Staubli VAL3: Motion.pjx

--- Motion.pjx ---
Parameters version=s8.15.3Cs9_BS3337 stackSize=200000 millimeterUnit=true
Program file=getMoveDone.pgx
Program file=home.pgx
Program file=moveToPoint.pgx
Program file=setSpeed.pgx
Data file=Motion.dtx
Library alias=io path=Disk://io/io.pjx autoload=true password=

--- Motion.dtx ---
public mdesc mNomSpeed = {accel=25, vel=20, decel=25, blend=off, leave=0, reach=0}
public mdesc mFine = {accel=10, vel=10, decel=10, blend=off, leave=0, reach=0}
public joint jHome
public tool tTool = {fatherId=flange[0]}

--- getMoveDone.pgx ---
public program getMoveDone(num& x_nResult)
  local num l_nT0
  local num l_nTimeout
//等待已下发的运动全部执行完，并等到机械臂停稳
//返回码 x_nResult：0=已停稳  1=指令执行完但 2s 内仍未停稳（残余抖动/受外力）
//依据：waitEndMove() 手册 10.6 第177页；isSettled() 手册 10.6 第178页
begin
  x_nResult=0

  //1) 取消上一条指令的混接，并等它执行完（手册 10.6，第177页）
  //   注意：waitEndMove 只等到"位置指令下发到位"，不等机械臂稳定
  waitEndMove()

  //2) 需要完全停稳时必须再用 isSettled()（手册 10.6，第178页）
  l_nTimeout=2
  if isSettled()==false
    l_nT0=clock()                                  //手册 5 章，第103页
    do
      delay(0.01)                                  //循环里必须让出 CPU
    until (isSettled()==true) or ((clock()-l_nT0)>=l_nTimeout)
    //超时不抛错：有的工位（打磨/压装）本来就有持续微振，交给调用方判断
    if isSettled()==false
      x_nResult=1
    endIf
  endIf
end

--- home.pgx ---
public program home(num& x_nResult)
  local num l_nMoveId
//关节运动(movej)回 Home 位 jHome，并等待到位/停稳
//返回码 x_nResult：0=已到 Home 并停稳  1=到点但仍有残余抖动  -2=jHome 超出软件限位
//依赖：Motion.dtx 的 jHome（当前是全 0 占位，示教后才是真实 Home）
begin
  x_nResult=0

  waitEndMove()

  //jHome 现在是全 0 占位，先判软件限位（bool isInRange(joint)，手册 9.2，第133页）；
  //不在限位内就直接返回错误，不要让控制器抛 runtime error
  if isInRange(jHome)==false
    x_nResult=-2
    return
  endIf

  //movej 的第一个参数必须用 joint 变量传入；写成 {0,0,0,0,0,0} 会被判为歧义表达式
  //（手册 10.6，第173页 movej 的 Example 有说明）
  l_nMoveId=movej(jHome,tTool,mFine)

  //move id 只能用 >= 判断，且完成判据是 +1（手册 10.4，第180页）
  wait(getMoveId()>=l_nMoveId+1)

  call getMoveDone(x_nResult)
end

--- moveToPoint.pgx ---
public program moveToPoint(point x_pTarget, tool x_tTool, mdesc x_mDesc, num& x_nResult)
  local num l_nMoveId
//直线运动(movel)到点位，并等待到位/停稳
//用法：call mot:moveToPoint(pPick, mot:tTool, mot:mNomSpeed, nResult)
//      要精定位时把第 3 个参数换成 mot:mFine
//返回码 x_nResult：0=已到位并停稳  1=指令执行完但仍有残余抖动（见 getMoveDone）  2=运动被中断
//点位由调用方传入（本库不放占位点位，见 Motion.dtx 注释）
begin
  x_nResult=0

  //0) 先把已下发的运动执行完，避免上一条指令的混接影响本次到位判断
  waitEndMove()

  //1) 下发直线运动，返回本次 move id（手册 10.6，第174页 num movel(point,tool,mdesc)）
  l_nMoveId=movel(x_pTarget,x_tTool,x_mDesc)

  //2) 等这条指令走过终点。move id 的整数部分是"正在执行的指令号"，
  //   指令刚下发时 getMoveId() 已经是 l_nMoveId.x，所以 >=l_nMoveId 会立刻成立；
  //   正确判据是 >=l_nMoveId+1（手册 10.4 第180页：waitEndMove 后 id = 最后一条 +1）
  wait(getMoveId()>=l_nMoveId+1)

  //3) 等机械臂真正停稳（waitEndMove 只等到指令执行完，不等稳定）
  call getMoveDone(x_nResult)
end

--- setSpeed.pgx ---
public program setSpeed(num x_nPercent, num& x_nResult)
  local mdesc l_mSpeed
  local num l_nAccel
//按百分比改 Motion.dtx 的 mNomSpeed（后续所有用 mNomSpeed 的运动都受影响）
//用法：call mot:setSpeed(50, nResult)   // 50%
//返回码 x_nResult：0=正常  -1=百分比越界（合法 1..100）
//字段含义见手册 10.5（第172页）：vel/accel/decel 均为额定值的百分比
begin
  x_nResult=0

  if (x_nPercent<1) or (x_nPercent>100)
    x_nResult=-1
    return
  endIf

  //先拷到局部 mdesc 再改字段，再整体写回（与参考工程 usrapp_dr/Move/setSpeed.pgx 同一写法）
  l_mSpeed=mNomSpeed
  l_mSpeed.vel=x_nPercent
  //加减速按速度平方折算，低速时加减速也小，避免小速度大加速度造成抖动
  l_nAccel=(x_nPercent*x_nPercent)/100
  l_mSpeed.accel=l_nAccel
  l_mSpeed.decel=l_nAccel
  //不在中间点混接，保证每条运动都精确到位（blend 取值 off/joint/Cartesian）
  l_mSpeed.blend=off
  l_mSpeed.leave=0
  l_mSpeed.reach=0

  mNomSpeed=l_mSpeed
end
